{attribute 'qualified_only'}
{attribute 'strict'}
TYPE E_ExTime :
(
	eCIP := 0,
	eWater,
	eProduct,
	eLine,
	eLineStby
);
END_TYPE

(* stored: Version 1.1.0.1, ProductVersion 3.1.4024.15
   DUT E_ExTime: Id {faf9b352-58b3-4d93-9c1c-ab4ea5941276} *)
